Fanuc KAREL source: ka00080.KL

-- PROVISIONAL review KL for V770-1; original PC SHA256 01218a3052bfc73d5a9bca4f060557c23944e4d7c2d9962e2dc68d59fbfc6b43
-- Incomplete behavior may be omitted. Consult companion uncertainty JSON. Do not deploy.
PROGRAM KA00080
%NOLOCKGROUP
-- UNRESOLVED_DECL SRC type=000106
-- UNRESOLVED_DECL DST type=000199
BEGIN
  -- UNRESOLVED_PC offsets 5-20; opcodes 2E,22,32,35
  -- UNRESOLVED_PC offsets 25-45; opcodes 49,7E,4A
  -- UNRESOLVED_PC offsets 50-54; opcodes 7F
END KA00080
